(* IEC 61131-3 sources: llm-plc-st-eval/data/processed_definitivo/qwen2.5-coder_14b/I1/zero_shot, 3 files *)

(* ---- ejec_1.st ---- *)
FUNCTION_BLOCK FB_Semaforo
VAR_INPUT
    habilitado : BOOL; // Variable de entrada que indica si el semáforo está habilitado
END_VAR

VAR_OUTPUT
    luzV : BOOL; // Variable de salida para la luz verde
    luzA : BOOL; // Variable de salida para la luz amarilla
    luzR : BOOL; // Variable de salida para la luz roja
END_VAR

VAR
    estado : INT := 0; // Variable de estado para controlar la secuencia del semáforo
    timer : TON; // Timer para controlar los tiempos de cada estado
    intermitente : BOOL := FALSE; // Variable para controlar el estado intermitente de la luz amarilla
END_VAR

// Inicialización del timer
timer(IN := TRUE, PT := T#20S);

// Máquina de estados
CASE estado OF
    0: // Estado verde
        luzV := TRUE;
        luzA := FALSE;
        luzR := FALSE;
        IF habilitado THEN
            IF timer.Q THEN
                timer(PT := T#4S); // Cambiar a amarillo después de 20 segundos
                estado := 1;
            END_IF
        ELSE
            estado := 3; // Cambiar a estado intermitente si habilitado se desactiva
        END_IF

    1: // Estado amarillo
        luzV := FALSE;
        luzA := TRUE;
        luzR := FALSE;
        IF habilitado THEN
            IF timer.Q THEN
                timer(PT := T#15S); // Cambiar a rojo después de 4 segundos
                estado := 2;
            END_IF
        ELSE
            estado := 3; // Cambiar a estado intermitente si habilitado se desactiva
        END_IF

    2: // Estado rojo
        luzV := FALSE;
        luzA := FALSE;
        luzR := TRUE;
        IF habilitado THEN
            IF timer.Q THEN
                timer(PT := T#20S); // Cambiar a verde después de 15 segundos
                estado := 0;
            END_IF
        ELSE
            estado := 3; // Cambiar a estado intermitente si habilitado se desactiva
        END_IF

    3: // Estado intermitente
        luzV := FALSE;
        luzA := intermitente;
        luzR := FALSE;
        IF habilitado THEN
            estado := 0; // Reiniciar la secuencia si habilitado se activa
        ELSE
            intermitente := NOT intermitente; // Cambiar el estado de intermitencia cada segundo
            timer(PT := T#1S); // Reiniciar el timer para el siguiente cambio de estado
        END_IF
END_CASE

(* ---- ejec_2.st ---- *)
FUNCTION_BLOCK FB_Semaforo
VAR_INPUT
    habilitado : BOOL; // Variable de entrada que indica si el semáforo está habilitado
END_VAR

VAR_OUTPUT
    luzV : BOOL; // Salida para la luz verde
    luzA : BOOL; // Salida para la luz amarilla
    luzR : BOOL; // Salida para la luz roja
END_VAR

VAR
    estado : INT := 0; // Variable de estado para controlar la secuencia
    contador : TON; // Contador de tiempo
    intermitente : BOOL := FALSE; // Variable para controlar el estado intermitente
END_VAR

// Inicialización del contador de tiempo
contador(IN := FALSE, PT := T#1S);

// Lógica del semáforo
CASE estado OF
    0: // Estado verde
        IF habilitado THEN
            luzV := TRUE;
            luzA := FALSE;
            luzR := FALSE;
            contador(IN := TRUE, PT := T#20S);
            IF contador.Q THEN
                estado := 1;
            END_IF;
        ELSE
            estado := 3; // Cambia a estado intermitente
        END_IF;

    1: // Estado amarillo
        IF habilitado THEN
            luzV := FALSE;
            luzA := TRUE;
            luzR := FALSE;
            contador(IN := TRUE, PT := T#4S);
            IF contador.Q THEN
                estado := 2;
            END_IF;
        ELSE
            estado := 3; // Cambia a estado intermitente
        END_IF;

    2: // Estado rojo
        IF habilitado THEN
            luzV := FALSE;
            luzA := FALSE;
            luzR := TRUE;
            contador(IN := TRUE, PT := T#15S);
            IF contador.Q THEN
                estado := 0;
            END_IF;
        ELSE
            estado := 3; // Cambia a estado intermitente
        END_IF;

    3: // Estado intermitente
        luzV := FALSE;
        luzA := intermitente;
        luzR := FALSE;
        contador(IN := TRUE, PT := T#1S);
        IF contador.Q THEN
            intermitente := NOT intermitente; // Cambia el estado intermitente
            contador(IN := FALSE); // Reinicia el contador
            IF habilitado THEN
                estado := 0; // Vuelve al estado verde si se habilita nuevamente
            END_IF;
        END_IF;

END_CASE

(* ---- ejec_3.st ---- *)
FUNCTION_BLOCK FB_Semaforo
VAR_INPUT
    habilitado : BOOL; // Entrada que habilita o deshabilita el semáforo
END_VAR

VAR_OUTPUT
    luzV : BOOL; // Salida para la luz verde
    luzA : BOOL; // Salida para la luz amarilla
    luzR : BOOL; // Salida para la luz roja
END_VAR

VAR
    estado : INT := 0; // Variable de estado para el semáforo
    timer : TON; // Timer para controlar los tiempos
    tiempoVerde : TIME := T#20S; // Tiempo verde
    tiempoAmarillo : TIME := T#4S; // Tiempo amarillo
    tiempoRojo : TIME := T#15S; // Tiempo rojo
    tiempoAmarilloIntermitente : TIME := T#1S; // Tiempo amarillo intermitente
    contadorAmarilloIntermitente : INT := 0; // Contador para el amarillo intermitente
END_VAR

// Inicialización del timer
timer(IN := FALSE, PT := tiempoVerde);

// Máquina de estados
CASE estado OF
    0: // Estado verde
        luzV := TRUE;
        luzA := FALSE;
        luzR := FALSE;
        IF habilitado THEN
            timer(IN := TRUE);
            IF timer.Q THEN
                timer(IN := FALSE);
                estado := 1; // Cambiar a estado amarillo
            END_IF
        ELSE
            estado := 3; // Cambiar a estado amarillo intermitente
        END_IF

    1: // Estado amarillo
        luzV := FALSE;
        luzA := TRUE;
        luzR := FALSE;
        IF habilitado THEN
            timer(IN := TRUE, PT := tiempoAmarillo);
            IF timer.Q THEN
                timer(IN := FALSE);
                estado := 2; // Cambiar a estado rojo
            END_IF
        ELSE
            estado := 3; // Cambiar a estado amarillo intermitente
        END_IF

    2: // Estado rojo
        luzV := FALSE;
        luzA := FALSE;
        luzR := TRUE;
        IF habilitado THEN
            timer(IN := TRUE, PT := tiempoRojo);
            IF timer.Q THEN
                timer(IN := FALSE);
                estado := 0; // Cambiar a estado verde
            END_IF
        ELSE
            estado := 3; // Cambiar a estado amarillo intermitente
        END_IF

    3: // Estado amarillo intermitente
        luzV := FALSE;
        luzA := contadorAmarilloIntermitente MOD 2 = 0;
        luzR := FALSE;
        IF habilitado THEN
            estado := 0; // Reiniciar a estado verde
        ELSE
            contadorAmarilloIntermitente := contadorAmarilloIntermitente + 1;
            timer(IN := TRUE, PT := tiempoAmarilloIntermitente);
        END_IF
END_CASE
